PROGRAM prg_LightTower
VAR_INPUT
	bBuzzerBypass: BOOL;
END_VAR
VAR

	ton_Blink				: TON;
	ton_Buzzer				: TON;
	t_Buzzer				: TIME:=T#2S;
	t_BuzzerShort			: TIME:=T#0.5S;
	t_BuzzerErrorDelay		: TIME:=T#10S;
	t_BuzzerWarningDelay	: TIME:=T#30S;
	//eLightTowerState_Last	: E_LightTowerState;
	bBuzzerMuteMemo: BOOL;	
	ton_MuteBuzzer: TON;
	ton_NoMessage: TON;
	ton_BuzzerLongTimeOn: TON;
END_VAR

VAR_OUTPUT
	qLedGreen	: BOOL;
	qLedYellow	: BOOL;
	qLedRed		: BOOL;
	qBuzzer		: BOOL;	
END_VAR

// Interface
(*
q_EL[1].ch1:=qLedGreen;
q_EL[1].ch2:=qLedYellow;
q_EL[1].ch3:=qLedRed;
q_EL[1].ch4:=qBuzzer;
*)
//.....................
(*
TYPE E_LightTowerState :
(
	eLightsOff := 0,
	eRed,				//Error
	eYellow,			//Pause
	eGreen,				//Run
	eGreenYellowBlink	//Run and warning
);
END_TYPE
*)
act_Operation();
ton_Blink(IN:=NOT ton_Blink.Q);
CASE eLightTowerState OF
	eLightsOff:;
		qLedGreen	:=FALSE;
		qLedYellow	:=FALSE;
		qLedRed		:=FALSE;
		eBuzzerMode:=eBuzzerOff;	
		
	eGreen:;
		qLedGreen	:=TRUE;
		qLedYellow	:=FALSE;
		qLedRed		:=FALSE;
		eBuzzerMode:=eBuzzerOff;	
		
	eGreen_YellowBlink:;
		qLedGreen	:=TRUE;
		qLedYellow	:=TRUE;
		qLedRed		:=FALSE;
		IF bBuzzerMuteMemo THEN;
			eBuzzerMode:=eBuzzerOff;
		ELSE
			eBuzzerMode:=eBuzzerWarning;
		END_IF
		ton_Blink.PT:=T#1S;
		IF ton_Blink.ET>T#0.5S THEN; qLedYellow:=FALSE; ELSE;qLedGreen:=FALSE; END_IF	
		
	eGreenBlink:;
		qLedGreen	:=TRUE;
		qLedYellow	:=FALSE;
		qLedRed		:=FALSE;
		eBuzzerMode:=eBuzzerOff;		
		ton_Blink.PT:=T#1S;
		IF ton_Blink.ET>T#0.5S THEN; qLedGreen:=FALSE; END_IF	

	eGreenBlink_YellowBlink:;
		qLedGreen	:=TRUE;
		qLedYellow	:=TRUE;
		qLedRed		:=FALSE;
		IF bBuzzerMuteMemo THEN;
			eBuzzerMode:=eBuzzerOff;
		ELSE
			eBuzzerMode:=eBuzzerWarning;
		END_IF
		ton_Blink.PT:=T#1S;
		IF ton_Blink.ET>T#0.5S THEN; qLedYellow:=FALSE; ELSE;qLedGreen:=FALSE; END_IF

	eGreenBlink_RedBlink:;
		qLedGreen	:=TRUE;
		qLedYellow	:=FALSE;
		qLedRed		:=TRUE;
		IF bBuzzerMuteMemo THEN;
			eBuzzerMode:=eBuzzerOff;
		ELSE
			eBuzzerMode:=eBuzzerError;
		END_IF
		ton_Blink.PT:=T#1S;
		IF ton_Blink.ET>T#0.5S THEN; qLedRed:=FALSE; ELSE;qLedGreen:=FALSE; END_IF
		
	eYellow:;
		qLedGreen	:=FALSE;
		qLedYellow	:=TRUE;
		qLedRed		:=FALSE;
		eBuzzerMode:=eBuzzerOff;	
		
	eRed:;
		qLedGreen	:=FALSE;
		qLedYellow	:=FALSE;
		qLedRed		:=TRUE;
		IF bBuzzerMuteMemo THEN;
			eBuzzerMode:=eBuzzerOff;
		ELSE
			eBuzzerMode:=eBuzzerError;
		END_IF
END_CASE

ton_NoMessage(PT:=T#5S,IN:=bBuzzerMuteMemo AND iActErrors=0 AND iActWarning=0);

IF (stOpMain.bSetPlay
	(*OR stOpLoad.bSetPlay
	OR stOpUnload.bSetPlay
	OR stOpManip.bSetPlay
	OR stOpHMI.bSetPlay
	OR prg_Call_OpMode.fbModeIndex.rt_Play.Q
	OR prg_Call_OpMode.fbModeLoad.rt_Play.Q
	OR prg_Call_OpMode.fbModeUnload.rt_Play.Q
	OR prg_Call_OpMode.fbModeManip.rt_Play.Q*)
	OR ton_NoMessage.Q	
)
THEN;
	ton_MuteBuzzer.IN:=TRUE;
END_IF
IF ton_MuteBuzzer.IN THEN;
	bBuzzerMuteMemo:=FALSE;
END_IF
ton_MuteBuzzer(PT:=T#1S);
IF ton_MuteBuzzer.Q THEN
	ton_MuteBuzzer.IN:=FALSE;
END_IF
IF prg_Messages.ResetErrors OR ton_BuzzerLongTimeOn.Q THEN;// iActErrors=0 AND iActWarning=0
	bBuzzerMuteMemo:=TRUE;
END_IF
ton_BuzzerLongTimeOn(PT:=T#30M,IN:=eBuzzerMode<>eBuzzerOff);

(*
TYPE E_BuzzerMode :
(
	eBuzzerOff := 0,
	eBuzzerError,		//Short Delay Off
	eBuzzerWarning		//Long Delay Off
);
END_TYPE
*)

IF NOT bBuzzerBypass THEN
	ton_Buzzer();
	CASE eBuzzerMode OF
		eBuzzerOff :;
			qBuzzer:=FALSE;
			
			ton_Buzzer.IN:=FALSE;
		eBuzzerError:;			//Short Delay Off
			qBuzzer:=TRUE;
			ton_Buzzer.PT:=t_BuzzerErrorDelay;
			ton_Buzzer.IN:=NOT ton_Buzzer.Q;
			IF ton_Buzzer.ET>t_Buzzer THEN; qBuzzer:=FALSE; END_IF
		eBuzzerWarning:;		//Long Delay Off
			qBuzzer:=TRUE;
			ton_Buzzer.PT:=t_BuzzerWarningDelay;
			ton_Buzzer.IN:=NOT ton_Buzzer.Q;
			IF ton_Buzzer.ET>t_BuzzerShort THEN; qBuzzer:=FALSE; END_IF
	END_CASE	
ELSE
	qBuzzer:=FALSE;
END_IF

ACTION act_Operation:
IF 		stOpMain.iActOperation=E_OperationButtons.ePauseAll
	AND iActErrors<>0
	THEN;	
	eLightTowerState:=E_LightTowerState.eRed;
 						//7
ELSIF 	stOpMain.iActOperation=E_OperationButtons.ePauseAll
	AND iActErrors=0
	THEN;
	eLightTowerState:=E_LightTowerState.eYellow;					//6	
	
ELSIF 	stOpMain.iActOperation=E_OperationButtons.ePlayAll
	AND iActErrors=0
 	AND iActWarning<>0
	THEN;
	eLightTowerState:=E_LightTowerState.eGreenBlink_YellowBlink;	//4
		
ELSIF 	stOpMain.iActOperation=E_OperationButtons.ePlayAll
	AND iActErrors=0 
	AND iActWarning=0 
	THEN;
	eLightTowerState:=E_LightTowerState.eGreen;						//1
END_IF
END_ACTION

ACTION act_Operation_Multi:
IF 		stOpMain.iActOperation=E_OperationButtons.ePauseAll
	//AND stOpLoad.iActOperation=E_OperationButtons.ePauseAll
	//AND stOpUnload.iActOperation=E_OperationButtons.ePauseAll
	//AND stOpManip.iActOperation=E_OperationButtons.ePauseAll
	//AND stOpHMI.iActOperation=E_OperationButtons.ePauseAll
	AND iActErrors<>0
	THEN;	
	eLightTowerState:=E_LightTowerState.eRed;
 						//7
ELSIF 	stOpMain.iActOperation=E_OperationButtons.ePauseAll
	//AND stOpLoad.iActOperation=E_OperationButtons.ePauseAll
	//AND stOpUnload.iActOperation=E_OperationButtons.ePauseAll
	//AND stOpManip.iActOperation=E_OperationButtons.ePauseAll
	//AND stOpHMI.iActOperation=E_OperationButtons.ePauseAll
	AND iActErrors=0
	THEN;
	eLightTowerState:=E_LightTowerState.eYellow;					//6
	
ELSIF 	(stOpMain.iActOperation=E_OperationButtons.ePlayAll
	(*OR stOpLoad.iActOperation=E_OperationButtons.ePlayAll
	OR stOpUnload.iActOperation=E_OperationButtons.ePlayAll
	OR stOpManip.iActOperation=E_OperationButtons.ePlayAll
	OR stOpHMI.iActOperation=E_OperationButtons.ePlayAll*))
	AND iActErrors<>0 
	THEN;
	eLightTowerState:=E_LightTowerState.eGreenBlink_RedBlink;		//5
	
ELSIF 	(stOpMain.iActOperation=E_OperationButtons.ePlayAll
	(*OR stOpLoad.iActOperation=E_OperationButtons.ePlayAll
	OR stOpUnload.iActOperation=E_OperationButtons.ePlayAll
	OR stOpManip.iActOperation=E_OperationButtons.ePlayAll
	OR stOpHMI.iActOperation=E_OperationButtons.ePlayAll*))
	AND iActErrors=0
 	AND iActWarning<>0
	THEN;
	eLightTowerState:=E_LightTowerState.eGreenBlink_YellowBlink;	//4
	
ELSIF  	(stOpMain.iActOperation=E_OperationButtons.ePlayAll
	(*OR stOpLoad.iActOperation=E_OperationButtons.ePlayAll
	OR stOpUnload.iActOperation=E_OperationButtons.ePlayAll
	OR stOpManip.iActOperation=E_OperationButtons.ePlayAll
	OR stOpHMI.iActOperation=E_OperationButtons.ePlayAll*))
	AND  (stOpMain.iActOperation=E_OperationButtons.ePauseAll
	(*OR stOpLoad.iActOperation=E_OperationButtons.ePauseAll
	OR stOpUnload.iActOperation=E_OperationButtons.ePauseAll
	OR stOpManip.iActOperation=E_OperationButtons.ePauseAll
	OR stOpHMI.iActOperation=E_OperationButtons.ePauseAll*))	
	AND iActErrors=0
 	AND iActWarning=0
	THEN;
	eLightTowerState:=E_LightTowerState.eGreenBlink;				//3
	
ELSIF 	stOpMain.iActOperation=E_OperationButtons.ePlayAll
	(*AND stOpLoad.iActOperation=E_OperationButtons.ePlayAll
	AND stOpUnload.iActOperation=E_OperationButtons.ePlayAll
	AND stOpManip.iActOperation=E_OperationButtons.ePlayAll
	AND stOpHMI.iActOperation=E_OperationButtons.ePlayAll*)
	AND iActErrors=0 
	AND iActWarning<>0
	THEN;
	eLightTowerState:=E_LightTowerState.eGreen_YellowBlink;			//2
	
ELSIF 	stOpMain.iActOperation=E_OperationButtons.ePlayAll
	(*AND stOpLoad.iActOperation=E_OperationButtons.ePlayAll
	AND stOpUnload.iActOperation=E_OperationButtons.ePlayAll
	AND stOpManip.iActOperation=E_OperationButtons.ePlayAll
	AND stOpHMI.iActOperation=E_OperationButtons.ePlayAll*)
	AND iActErrors=0 
	AND iActWarning=0 
	THEN;
	eLightTowerState:=E_LightTowerState.eGreen;						//1
END_IF
END_ACTION

END_PROGRAM

(* stored: Version 1.1.0.1, ProductVersion 3.1.4024.13
   POU prg_LightTower: Id {f02147ec-0518-45ea-a1e9-951e541f9e2a}, SpecialFunc None
   Action act_Operation: Id {8d6c7f2a-28a2-4a68-b801-679d7d75691a}
   Action act_Operation_Multi: Id {bd77fe55-28e8-42fd-84e0-4c32f2e825d2} *)
